// HAL boundary for one analog output channel. The composition root maps the
// raw process value from here; identity is injected separately (S10.2.1).
TYPE ST_AnalogOutputHal :
STRUCT
    Raw : LREAL;
END_STRUCT
END_TYPE

(* stored: Version 1.1.0.1, ProductVersion 3.1.4024.12
   DUT ST_AnalogOutputHal: Id {3bbd4f76-bda6-48a1-ac31-246cda7a20ee} *)
